(* IEC 61131-3 sources: sis-interlock-demo/tests/POUs/Helpers/FB_VotingRig, 8 files *)

(* ---- FB_VotingRig.decl.st ---- *)
// Назначение: стенд тестов FB_Voting: подменное время (старт LTIME#1H), журнал событий и группа
//             голосования; тест пишет входы стенда и вызывает Cycle/Step/Run.
// Автор:      kr0nsch
// Версия:     0.1.0
// Документ:   docs/DESIGN.md, раздел «12.3 Граничные случаи (вручную, команда A)»
// ВНИМАНИЕ:   код демонстрационный и не предназначен для систем безопасности. Реальная ПАЗ
//             требует определения SIL, сертифицированных аппаратных и программных средств
//             и валидации по ГОСТ Р МЭК 61511.
FUNCTION_BLOCK FB_VotingRig
VAR_INPUT
    stIn          : ST_VoteIn;          // сигналы каналов
    stCmd         : ST_VoteCmd;         // запросы байпаса
    stCfg         : ST_VotingCfg;       // конфигурация группы
    xBypassPermit : BOOL := TRUE;       // ключ разрешения байпасов
    uiCause       : UINT := 7;          // номер причины в событиях
END_VAR
VAR
    fbTime : PL.FB_FakeTime;            // подменное время
    fbLog  : FB_SisTestLog;             // журнал событий
    fbVote : FB_Voting;                 // ФБ под тестом
END_VAR

(* ---- BypassOf.method.decl.st ---- *)
// Код состояния байпаса канала (TO_INT(E_BypassState))
METHOD BypassOf : INT
VAR_INPUT
    uiCh : UINT;   // номер канала
END_VAR

(* ---- Run.method.decl.st ---- *)
// Шаги tStep до tDuration (последний — остаток), вызов после каждого шага; не больше 1500 шагов
METHOD Run
VAR_INPUT
    tDuration : TIME;   // сколько времени пройти
    tStep     : TIME;   // шаг
END_VAR
VAR
    tLeft  : TIME;      // осталось
    tNow   : TIME;      // этот шаг
    uiIter : UINT;      // шагов сделано
END_VAR

(* ---- SetAi.method.decl.st ---- *)
// Значения аналоговых каналов 1..3, все достоверны
METHOD SetAi
VAR_INPUT
    r1 : REAL;   // канал 1, инж. ед.
    r2 : REAL;   // канал 2, инж. ед.
    r3 : REAL;   // канал 3, инж. ед.
END_VAR

(* ---- SetDi.method.decl.st ---- *)
// Значения дискретных каналов 1..3, линия у всех исправна
METHOD SetDi
VAR_INPUT
    x1 : BOOL;   // канал 1
    x2 : BOOL;   // канал 2
    x3 : BOOL;   // канал 3
END_VAR

(* ---- SetNow.method.decl.st ---- *)
// Установить подменное время (в том числе назад)
METHOD SetNow
VAR_INPUT
    ltValue : LTIME;   // новое время
END_VAR

(* ---- StateOf.method.decl.st ---- *)
// Код состояния канала (TO_INT(E_ChannelState))
METHOD StateOf : INT
VAR_INPUT
    uiCh : UINT;   // номер канала
END_VAR

(* ---- Step.method.decl.st ---- *)
// Продвинуть время на шаг и вызвать FB_Voting
METHOD Step
VAR_INPUT
    tStep : TIME;   // шаг времени
END_VAR
